// TIA Portal V20 export
Screen "HTML_VIEW"  1276x673
  ScreenItem "Title_ScreenOverview_X390_Y2" at 390,2 size 500x30  Type=HmiTextBox
  ScreenItem "Line_Header_X0_Y64" at 0,64 size 1276x0  Type=HmiLine
  ScreenItem "Text_DeviceAdress" at 390,36 size 150x25  Type=HmiTextBox
  ScreenItem "EA-Field_DeviceAdress" at 540,36 size 350x25  Type=HmiIOField
  ScreenItem "permanentareaborderrectangle" at 0,0 size 0x0  Type=HmiRectangle
  ScreenItem "网络控件_1" at 0,68 size 1280x586  Type=HmiWebControl
  ScreenItem "Button_Back" at 2,2 size 90x60  Type=HmiButton
